ABB RAPID module: MainProgram.mod

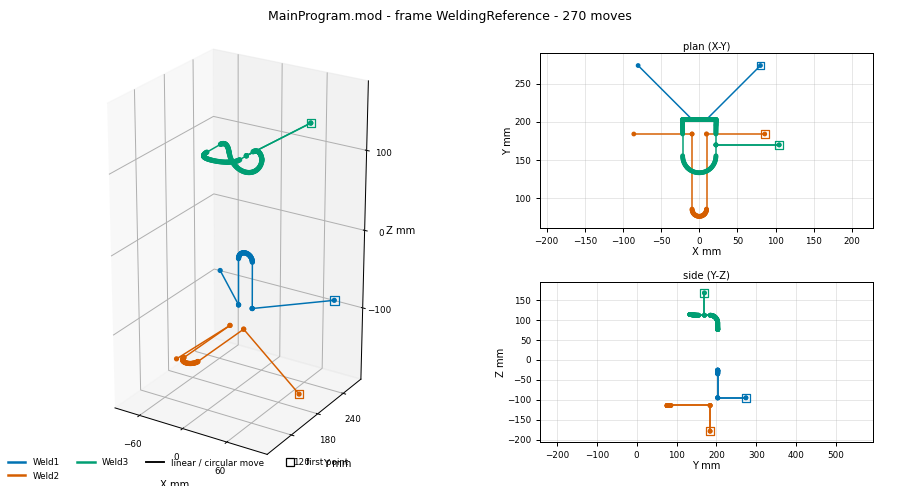
[picture p0: tool path of MainProgram.mod in frame WeldingReference, 270 of 274 moves have a stored position in this frame; points joined in program order, loops and branches not executed]
%%%
  VERSION:1
  LANGUAGE:ENGLISH
%%%
MODULE MOD_MainProgram

    ! -------------------------------
    ! Define customized variables here
    ! ...

	! Tool variables:
	PERS tooldata Weldgun := [TRUE,[[-4.000,0.000,371.300],[0.92387953,0.00000000,0.38268343,0.00000001]],[1,[0,0,20],[1,0,0,0],0,0,0.005]];

	! Reference variables:
	PERS wobjdata WeldingReference := [FALSE, TRUE, "", [[0,0,0],[1,0,0,0]],[[907.213,-302.346,276.168],[0.70442562,0.70442562,-0.06151869,-0.06151869]]];

	PROC GoHome()
		ConfJ \On;
		ConfL \Off;
		MoveAbsJ [[-0.000000,-14.941300,9.781060,0.000000,57.564300,-0.000000],[9E+09,9E+09,9E+09,9E+09,9E+09,9E+09]],v500,z1,Weldgun \WObj:=WeldingReference;
	ENDPROC

	PROC Weld1()
		ConfJ \On;
		ConfL \Off;
		WeldingReference := [FALSE, TRUE, "", [[0,0,0],[1,0,0,0]],[[907.213,-302.346,276.168],[0.70442562,0.70442562,-0.06151869,-0.06151869]]];
		Weldgun := [TRUE,[[-4.000,0.000,371.300],[0.92387953,0.00000000,0.38268343,0.00000001]],[1,[0,0,20],[1,0,0,0],0,0,0.005]];
		! show Weld gun
		MoveAbsJ [[-12.555800,6.650190,11.177100,0.026927,72.173900,-2.607590],[9E+09,9E+09,9E+09,9E+09,9E+09,9E+09]],v1000,z1,Weldgun \WObj:=WeldingReference;
		SetRPM 70.0;
		MoveL [[80.178,273.912,-94.776],[0.27080492,-0.27039115,-0.65336714,0.65319576],[-1,0,-1,0],[9E+09,9E+09,9E+09,9E+09,9E+09,9E+09]],[16.67,500,5000,1000],z1,Weldgun \WObj:=WeldingReference;
		MoveL [[9.468,203.201,-94.776],[0.27080492,-0.27039115,-0.65336714,0.65319576],[-1,0,-1,0],[9E+09,9E+09,9E+09,9E+09,9E+09,9E+09]],[16.67,500,5000,1000],z1,Weldgun \WObj:=WeldingReference;
		GunOn;
		MoveL [[9.468,203.201,-94.776],[0.27080492,-0.27039115,-0.65336714,0.65319576],[-1,0,-1,0],[9E+09,9E+09,9E+09,9E+09,9E+09,9E+09]],[16.67,500,5000,1000],z1,Weldgun \WObj:=WeldingReference;
		MoveL [[9.521,203.201,-94.770],[0.27059813,-0.27059797,-0.65328151,0.65328145],[-1,0,-1,0],[9E+09,9E+09,9E+09,9E+09,9E+09,9E+09]],[16.67,500,5000,1000],z1,Weldgun \WObj:=WeldingReference;
		MoveL [[9.521,203.201,-34.925],[0.26109596,-0.28004323,-0.64928868,0.65713689],[-1,-1,-1,0],[9E+09,9E+09,9E+09,9E+09,9E+09,9E+09]],[16.67,500,5000,1000],z1,Weldgun \WObj:=WeldingReference;
		MoveL [[9.489,203.201,-34.145],[0.23425026,-0.30675221,-0.65944853,0.64510273],[-1,-1,0,0],[9E+09,9E+09,9E+09,9E+09,9E+09,9E+09]],[16.67,500,5000,1000],z1,Weldgun \WObj:=WeldingReference;
		MoveL [[9.394,203.201,-33.370],[0.20701375,-0.33294335,-0.66849979,0.63198265],[-1,-1,0,0],[9E+09,9E+09,9E+09,9E+09,9E+09,9E+09]],[16.67,500,5000,1000],z1,Weldgun \WObj:=WeldingReference;
		MoveL [[9.235,203.201,-32.605],[0.17943264,-0.35858122,-0.67642029,0.61780177],[-1,-1,0,0],[9E+09,9E+09,9E+09,9E+09,9E+09,9E+09]],[16.67,500,5000,1000],z1,Weldgun \WObj:=WeldingReference;
		MoveL [[9.014,203.201,-31.857],[0.15154219,-0.38361099,-0.68321444,0.60257415],[-1,-1,0,0],[9E+09,9E+09,9E+09,9E+09,9E+09,9E+09]],[16.67,500,5000,1000],z1,Weldgun \WObj:=WeldingReference;
		MoveL [[8.732,203.201,-31.128],[0.12340353,-0.40798899,-0.68885701,0.58633828],[-1,-1,0,0],[9E+09,9E+09,9E+09,9E+09,9E+09,9E+09]],[16.67,500,5000,1000],z1,Weldgun \WObj:=WeldingReference;
		MoveL [[8.391,203.201,-30.426],[0.09505233,-0.43169103,-0.69333556,0.56911660],[-1,-1,0,0],[9E+09,9E+09,9E+09,9E+09,9E+09,9E+09]],[16.67,500,5000,1000],z1,Weldgun \WObj:=WeldingReference;
		MoveL [[7.994,203.201,-29.753],[0.06655006,-0.45466761,-0.69664493,0.55093947],[-1,-1,0,0],[9E+09,9E+09,9E+09,9E+09,9E+09,9E+09]],[16.67,500,5000,1000],z1,Weldgun \WObj:=WeldingReference;
		MoveL [[7.544,203.201,-29.116],[0.03792629,-0.47687790,-0.69878733,0.53183205],[-1,-1,0,0],[9E+09,9E+09,9E+09,9E+09,9E+09,9E+09]],[16.67,500,5000,1000],z1,Weldgun \WObj:=WeldingReference;
		MoveL [[7.042,203.201,-28.517],[0.01240330,-0.49395227,-0.70281556,0.51176909],[-1,-1,0,0],[9E+09,9E+09,9E+09,9E+09,9E+09,9E+09]],[16.67,500,5000,1000],z1,Weldgun \WObj:=WeldingReference;
		MoveL [[6.733,203.201,-28.192],[0.00416831,0.50587340,0.70291668,-0.49998286],[-1,-1,0,0],[9E+09,9E+09,9E+09,9E+09,9E+09,9E+09]],[16.67,500,5000,1000],z1,Weldgun \WObj:=WeldingReference;
		MoveL [[6.408,203.201,-27.883],[0.02374061,0.52184249,0.69941540,-0.48778571],[-1,-1,0,0],[9E+09,9E+09,9E+09,9E+09,9E+09,9E+09]],[16.67,500,5000,1000],z1,Weldgun \WObj:=WeldingReference;
		MoveL [[5.809,203.201,-27.381],[0.05240062,0.54140968,0.69785181,-0.46597487],[-1,-1,0,0],[9E+09,9E+09,9E+09,9E+09,9E+09,9E+09]],[16.67,500,5000,1000],z1,Weldgun \WObj:=WeldingReference;
		MoveL [[5.172,203.201,-26.930],[0.08097272,0.56005587,0.69511960,-0.44338425],[-1,-1,0,0],[9E+09,9E+09,9E+09,9E+09,9E+09,9E+09]],[16.67,500,5000,1000],z1,Weldgun \WObj:=WeldingReference;
		MoveL [[4.499,203.201,-26.534],[0.10940637,0.57776774,0.69121158,-0.42004909],[-1,-1,0,0],[9E+09,9E+09,9E+09,9E+09,9E+09,9E+09]],[16.67,500,5000,1000],z1,Weldgun \WObj:=WeldingReference;
		MoveL [[3.797,203.201,-26.193],[0.13765258,0.59450380,0.68614585,-0.39600615],[-1,-1,0,0],[9E+09,9E+09,9E+09,9E+09,9E+09,9E+09]],[16.67,500,5000,1000],z1,Weldgun \WObj:=WeldingReference;
		MoveL [[3.068,203.201,-25.912],[0.16567219,0.61024237,0.67992465,-0.37129428],[-1,-1,0,0],[9E+09,9E+09,9E+09,9E+09,9E+09,9E+09]],[16.67,500,5000,1000],z1,Weldgun \WObj:=WeldingReference;
		MoveL [[2.320,203.201,-25.690],[0.19341081,0.62495524,0.67255736,-0.34596213],[-1,-1,0,0],[9E+09,9E+09,9E+09,9E+09,9E+09,9E+09]],[16.67,500,5000,1000],z1,Weldgun \WObj:=WeldingReference;
		MoveL [[1.555,203.201,-25.531],[0.22082406,0.63861348,0.66406224,-0.32004826],[-1,-1,0,0],[9E+09,9E+09,9E+09,9E+09,9E+09,9E+09]],[16.67,500,5000,1000],z1,Weldgun \WObj:=WeldingReference;
		MoveL [[0.780,203.201,-25.436],[0.24786932,0.65119902,0.65444982,-0.29359169],[-1,-1,0,0],[9E+09,9E+09,9E+09,9E+09,9E+09,9E+09]],[16.67,500,5000,1000],z1,Weldgun \WObj:=WeldingReference;
		MoveL [[0.000,203.201,-25.404],[0.27449275,0.66268723,0.64373837,-0.26664635],[-1,-1,0,0],[9E+09,9E+09,9E+09,9E+09,9E+09,9E+09]],[16.67,500,5000,1000],z1,Weldgun \WObj:=WeldingReference;
		MoveL [[-0.780,203.201,-25.436],[0.30065949,0.67306272,0.63194229,-0.23924755],[-1,-1,0,0],[9E+09,9E+09,9E+09,9E+09,9E+09,9E+09]],[16.67,500,5000,1000],z1,Weldgun \WObj:=WeldingReference;
		MoveL [[-1.555,203.201,-25.531],[0.32631571,0.68230801,0.61908153,-0.21145189],[-1,0,1,0],[9E+09,9E+09,9E+09,9E+09,9E+09,9E+09]],[16.67,500,5000,1000],z1,Weldgun \WObj:=WeldingReference;
		MoveL [[-2.320,203.201,-25.690],[0.35142970,0.69040355,0.60518073,-0.18329319],[-1,0,1,0],[9E+09,9E+09,9E+09,9E+09,9E+09,9E+09]],[16.67,500,5000,1000],z1,Weldgun \WObj:=WeldingReference;
		MoveL [[-3.068,203.201,-25.912],[0.37594474,0.69734095,0.59026085,-0.15483308],[-1,0,1,0],[9E+09,9E+09,9E+09,9E+09,9E+09,9E+09]],[16.67,500,5000,1000],z1,Weldgun \WObj:=WeldingReference;
		MoveL [[-3.797,203.201,-26.193],[0.39983154,0.70309811,0.57435509,-0.12611111],[-1,0,1,0],[9E+09,9E+09,9E+09,9E+09,9E+09,9E+09]],[16.67,500,5000,1000],z1,Weldgun \WObj:=WeldingReference;
		MoveL [[-4.499,203.201,-26.534],[0.42304339,0.70768163,0.55747448,-0.09717615],[-1,0,1,0],[9E+09,9E+09,9E+09,9E+09,9E+09,9E+09]],[16.67,500,5000,1000],z1,Weldgun \WObj:=WeldingReference;
		MoveL [[-5.172,203.201,-26.930],[0.44554480,0.71107104,0.53966024,-0.06807809],[-1,0,1,0],[9E+09,9E+09,9E+09,9E+09,9E+09,9E+09]],[16.67,500,5000,1000],z1,Weldgun \WObj:=WeldingReference;
		MoveL [[-5.809,203.201,-27.381],[0.46730140,0.71326404,0.52093536,-0.03886082],[-1,0,1,0],[9E+09,9E+09,9E+09,9E+09,9E+09,9E+09]],[16.67,500,5000,1000],z1,Weldgun \WObj:=WeldingReference;
		MoveL [[-6.408,203.201,-27.883],[0.48819595,0.71113015,0.50576611,-0.01261974],[-1,0,1,0],[9E+09,9E+09,9E+09,9E+09,9E+09,9E+09]],[16.67,500,5000,1000],z1,Weldgun \WObj:=WeldingReference;
		MoveL [[-6.731,203.201,-28.191],[0.49992546,0.71126987,0.49411825,0.00410579],[-1,0,1,0],[9E+09,9E+09,9E+09,9E+09,9E+09,9E+09]],[16.67,500,5000,1000],z1,Weldgun \WObj:=WeldingReference;
		MoveL [[-7.042,203.201,-28.517],[0.51134749,0.71391546,0.47777457,0.02408169],[-1,0,1,0],[9E+09,9E+09,9E+09,9E+09,9E+09,9E+09]],[16.67,500,5000,1000],z1,Weldgun \WObj:=WeldingReference;
		MoveL [[-7.544,203.201,-29.116],[0.53050914,0.71232829,0.45640294,0.05333687],[-1,0,1,0],[9E+09,9E+09,9E+09,9E+09,9E+09,9E+09]],[16.67,500,5000,1000],z1,Weldgun \WObj:=WeldingReference;
		MoveL [[-7.994,203.201,-29.753],[0.54878026,0.70953905,0.43426730,0.08250137],[-1,0,1,0],[9E+09,9E+09,9E+09,9E+09,9E+09,9E+09]],[16.67,500,5000,1000],z1,Weldgun \WObj:=WeldingReference;
		MoveL [[-8.391,203.201,-30.426],[0.56612441,0.70556165,0.41139698,0.11152774],[-1,0,1,0],[9E+09,9E+09,9E+09,9E+09,9E+09,9E+09]],[16.67,500,5000,1000],z1,Weldgun \WObj:=WeldingReference;
		MoveL [[-8.732,203.201,-31.128],[0.58251728,0.70039316,0.38784300,0.14035973],[-1,0,1,0],[9E+09,9E+09,9E+09,9E+09,9E+09,9E+09]],[16.67,500,5000,1000],z1,Weldgun \WObj:=WeldingReference;
		MoveL [[-9.014,203.201,-31.857],[0.59792965,0.69404912,0.36363243,0.16895976],[-1,0,1,0],[9E+09,9E+09,9E+09,9E+09,9E+09,9E+09]],[16.67,500,5000,1000],z1,Weldgun \WObj:=WeldingReference;
		MoveL [[-9.235,203.201,-32.605],[0.61233261,0.68654186,0.33880881,0.19727554],[-1,0,1,0],[9E+09,9E+09,9E+09,9E+09,9E+09,9E+09]],[16.67,500,5000,1000],z1,Weldgun \WObj:=WeldingReference;
		MoveL [[-9.394,203.201,-33.370],[0.62571166,0.67787385,0.31341661,0.22525981],[-1,0,1,0],[9E+09,9E+09,9E+09,9E+09,9E+09,9E+09]],[16.67,500,5000,1000],z1,Weldgun \WObj:=WeldingReference;
		MoveL [[-9.489,203.201,-34.145],[0.63803534,0.66806855,0.28749564,0.25286671],[-1,0,1,0],[9E+09,9E+09,9E+09,9E+09,9E+09,9E+09]],[16.67,500,5000,1000],z1,Weldgun \WObj:=WeldingReference;
		MoveL [[-9.521,203.201,-34.925],[0.65328148,0.65328148,0.27059805,0.27059805],[-1,0,1,0],[9E+09,9E+09,9E+09,9E+09,9E+09,9E+09]],[16.67,500,5000,1000],z1,Weldgun \WObj:=WeldingReference;
		MoveL [[-9.521,203.201,-94.770],[0.65328148,0.65328148,0.27059805,0.27059805],[-1,0,1,0],[9E+09,9E+09,9E+09,9E+09,9E+09,9E+09]],[16.67,500,5000,1000],z1,Weldgun \WObj:=WeldingReference;
		MoveL [[-9.470,203.201,-94.776],[0.65328148,0.65328148,0.27059805,0.27059805],[-1,0,1,0],[9E+09,9E+09,9E+09,9E+09,9E+09,9E+09]],[16.67,500,5000,1000],z1,Weldgun \WObj:=WeldingReference;
		GunOff;
		MoveL [[-9.470,203.201,-94.776],[0.65328148,0.65328148,0.27059805,0.27059805],[-1,0,1,0],[9E+09,9E+09,9E+09,9E+09,9E+09,9E+09]],v1000,z1,Weldgun \WObj:=WeldingReference;
		MoveL [[-80.181,273.912,-94.776],[0.65328148,0.65328148,0.27059805,0.27059805],[-1,0,1,0],[9E+09,9E+09,9E+09,9E+09,9E+09,9E+09]],v1000,z1,Weldgun \WObj:=WeldingReference;
	ENDPROC

	PROC Weld2()
		ConfJ \On;
		ConfL \Off;
		WeldingReference := [FALSE, TRUE, "", [[0,0,0],[1,0,0,0]],[[907.213,-302.346,276.168],[0.70442562,0.70442562,-0.06151869,-0.06151869]]];
		Weldgun := [TRUE,[[-4.000,0.000,371.300],[0.92387953,0.00000000,0.38268343,0.00000001]],[1,[0,0,20],[1,0,0,0],0,0,0.005]];
		! show Weld gun
		MoveAbsJ [[14.847000,37.704900,12.622700,-66.388600,108.377000,54.200400],[9E+09,9E+09,9E+09,9E+09,9E+09,9E+09]],v1000,z1,Weldgun \WObj:=WeldingReference;
		SetRPM 70.0;
		MoveL [[85.827,184.150,-178.501],[0.00000000,-0.42074767,0.00000000,0.90717771],[0,-1,0,0],[9E+09,9E+09,9E+09,9E+09,9E+09,9E+09]],[16.67,500,5000,1000],z1,Weldgun \WObj:=WeldingReference;
		MoveL [[9.489,184.150,-113.907],[0.00000000,-0.42074767,0.00000000,0.90717771],[0,-1,0,0],[9E+09,9E+09,9E+09,9E+09,9E+09,9E+09]],[16.67,500,5000,1000],z1,Weldgun \WObj:=WeldingReference;
		GunOn;
		MoveL [[9.489,184.150,-113.907],[0.00000000,-0.42074767,0.00000000,0.90717771],[0,-1,0,0],[9E+09,9E+09,9E+09,9E+09,9E+09,9E+09]],[16.67,500,5000,1000],z1,Weldgun \WObj:=WeldingReference;
		MoveL [[9.489,85.725,-113.907],[0.01312106,-0.42070385,-0.00608599,0.90708273],[0,-1,0,0],[9E+09,9E+09,9E+09,9E+09,9E+09,9E+09]],[16.67,500,5000,1000],z1,Weldgun \WObj:=WeldingReference;
		MoveL [[9.457,84.942,-113.910],[0.05153547,-0.42042592,0.00808679,0.90582600],[0,-1,0,0],[9E+09,9E+09,9E+09,9E+09,9E+09,9E+09]],[16.67,500,5000,1000],z1,Weldgun \WObj:=WeldingReference;
		MoveL [[9.361,84.163,-113.917],[0.08985371,-0.41918442,0.02228324,0.90316897],[0,-1,0,0],[9E+09,9E+09,9E+09,9E+09,9E+09,9E+09]],[16.67,500,5000,1000],z1,Weldgun \WObj:=WeldingReference;
		MoveL [[9.202,83.396,-113.930],[0.12804465,-0.41698615,0.03650971,0.89910742],[0,-1,0,0],[9E+09,9E+09,9E+09,9E+09,9E+09,9E+09]],[16.67,500,5000,1000],z1,Weldgun \WObj:=WeldingReference;
		MoveL [[8.981,82.644,-113.948],[0.16597915,-0.41384219,0.05079357,0.89364735],[0,-1,0,0],[9E+09,9E+09,9E+09,9E+09,9E+09,9E+09]],[16.67,500,5000,1000],z1,Weldgun \WObj:=WeldingReference;
		MoveL [[8.700,81.913,-113.970],[0.20363787,-0.40977344,0.06511381,0.88677931],[0,-1,0,0],[9E+09,9E+09,9E+09,9E+09,9E+09,9E+09]],[16.67,500,5000,1000],z1,Weldgun \WObj:=WeldingReference;
		MoveL [[8.360,81.208,-113.995],[0.24095022,-0.40479903,0.07948489,0.87850037],[0,-1,0,0],[9E+09,9E+09,9E+09,9E+09,9E+09,9E+09]],[16.67,500,5000,1000],z1,Weldgun \WObj:=WeldingReference;
		MoveL [[7.963,80.534,-114.024],[0.27783978,-0.39894829,0.09389601,0.86880887],[0,-1,0,0],[9E+09,9E+09,9E+09,9E+09,9E+09,9E+09]],[16.67,500,5000,1000],z1,Weldgun \WObj:=WeldingReference;
		MoveL [[7.512,79.895,-114.054],[0.31416482,-0.39224451,0.10838187,0.85772844],[0,-1,0,0],[9E+09,9E+09,9E+09,9E+09,9E+09,9E+09]],[16.67,500,5000,1000],z1,Weldgun \WObj:=WeldingReference;
		MoveL [[7.009,79.295,-114.086],[0.34473394,-0.38397214,0.12525349,0.84736974],[0,-1,0,0],[9E+09,9E+09,9E+09,9E+09,9E+09,9E+09]],[16.67,500,5000,1000],z1,Weldgun \WObj:=WeldingReference;
		MoveL [[6.707,78.978,-114.104],[0.36453651,-0.37938408,0.13335075,0.83988001],[0,-1,0,0],[9E+09,9E+09,9E+09,9E+09,9E+09,9E+09]],[16.67,500,5000,1000],z1,Weldgun \WObj:=WeldingReference;
		MoveL [[6.391,78.676,-114.123],[0.38912980,-0.37541067,0.13918584,0.82962168],[0,-1,0,0],[9E+09,9E+09,9E+09,9E+09,9E+09,9E+09]],[16.67,500,5000,1000],z1,Weldgun \WObj:=WeldingReference;
		MoveL [[5.795,78.176,-114.154],[0.42321516,-0.36636835,0.15366636,0.81427871],[0,-1,0,0],[9E+09,9E+09,9E+09,9E+09,9E+09,9E+09]],[16.67,500,5000,1000],z1,Weldgun \WObj:=WeldingReference;
		MoveL [[5.160,77.727,-114.185],[0.45649477,-0.35666115,0.16813439,0.79758145],[0,-1,0,0],[9E+09,9E+09,9E+09,9E+09,9E+09,9E+09]],[16.67,500,5000,1000],z1,Weldgun \WObj:=WeldingReference;
		MoveL [[4.490,77.331,-114.213],[0.48887672,-0.34632893,0.18258429,0.77956321],[0,-1,0,0],[9E+09,9E+09,9E+09,9E+09,9E+09,9E+09]],[16.67,500,5000,1000],z1,Weldgun \WObj:=WeldingReference;
		MoveL [[3.790,76.991,-114.239],[0.52034210,-0.33543360,0.19697026,0.76021781],[0,-1,-1,0],[9E+09,9E+09,9E+09,9E+09,9E+09,9E+09]],[16.67,500,5000,1000],z1,Weldgun \WObj:=WeldingReference;
		MoveL [[3.063,76.710,-114.260],[0.55080992,-0.32401460,0.21128182,0.73958297],[0,-1,-1,0],[9E+09,9E+09,9E+09,9E+09,9E+09,9E+09]],[16.67,500,5000,1000],z1,Weldgun \WObj:=WeldingReference;
		MoveL [[2.316,76.490,-114.278],[0.58023779,-0.31212946,0.22547321,0.71767759],[0,-1,-1,0],[9E+09,9E+09,9E+09,9E+09,9E+09,9E+09]],[16.67,500,5000,1000],z1,Weldgun \WObj:=WeldingReference;
		MoveL [[1.553,76.331,-114.291],[0.60858630,-0.29982600,0.23951509,0.69452113],[0,-1,-1,0],[9E+09,9E+09,9E+09,9E+09,9E+09,9E+09]],[16.67,500,5000,1000],z1,Weldgun \WObj:=WeldingReference;
		MoveL [[0.779,76.236,-114.299],[0.63581862,-0.28715637,0.25336406,0.67013622],[0,-1,-1,0],[9E+09,9E+09,9E+09,9E+09,9E+09,9E+09]],[16.67,500,5000,1000],z1,Weldgun \WObj:=WeldingReference;
		MoveL [[0.000,76.204,-114.301],[0.66190027,-0.27416831,0.26698017,0.64454741],[0,-1,-1,0],[9E+09,9E+09,9E+09,9E+09,9E+09,9E+09]],[16.67,500,5000,1000],z1,Weldgun \WObj:=WeldingReference;
		MoveL [[-0.779,76.236,-114.299],[0.68679970,-0.26090700,0.28032057,0.61778159],[0,-1,-1,0],[9E+09,9E+09,9E+09,9E+09,9E+09,9E+09]],[16.67,500,5000,1000],z1,Weldgun \WObj:=WeldingReference;
		MoveL [[-1.553,76.331,-114.291],[0.71048565,-0.24741615,0.29333969,0.58987051],[0,-1,-1,0],[9E+09,9E+09,9E+09,9E+09,9E+09,9E+09]],[16.67,500,5000,1000],z1,Weldgun \WObj:=WeldingReference;
		MoveL [[-2.316,76.490,-114.278],[0.73293327,-0.23373805,0.30598954,0.56084377],[0,-1,-1,0],[9E+09,9E+09,9E+09,9E+09,9E+09,9E+09]],[16.67,500,5000,1000],z1,Weldgun \WObj:=WeldingReference;
		MoveL [[-3.063,76.710,-114.260],[0.75411156,-0.21990803,0.31822287,0.53074516],[0,-1,-1,0],[9E+09,9E+09,9E+09,9E+09,9E+09,9E+09]],[16.67,500,5000,1000],z1,Weldgun \WObj:=WeldingReference;
		MoveL [[-3.790,76.991,-114.239],[0.77400420,-0.20596628,0.32998612,0.49960440],[0,-1,-1,0],[9E+09,9E+09,9E+09,9E+09,9E+09,9E+09]],[16.67,500,5000,1000],z1,Weldgun \WObj:=WeldingReference;
		MoveL [[-4.490,77.331,-114.213],[0.79256096,-0.19192832,0.34123966,0.46751058],[0,-1,-1,0],[9E+09,9E+09,9E+09,9E+09,9E+09,9E+09]],[16.67,500,5000,1000],z1,Weldgun \WObj:=WeldingReference;
		MoveL [[-5.160,77.727,-114.185],[0.80978515,-0.17783865,0.35192282,0.43447872],[0,-1,-1,0],[9E+09,9E+09,9E+09,9E+09,9E+09,9E+09]],[16.67,500,5000,1000],z1,Weldgun \WObj:=WeldingReference;
		MoveL [[-5.795,78.176,-114.154],[0.82563537,-0.16370520,0.36199413,0.40060840],[0,-1,-1,0],[9E+09,9E+09,9E+09,9E+09,9E+09,9E+09]],[16.67,500,5000,1000],z1,Weldgun \WObj:=WeldingReference;
		MoveL [[-6.391,78.676,-114.123],[0.83783925,-0.14727053,0.37231303,0.37110616],[0,-1,-1,0],[9E+09,9E+09,9E+09,9E+09,9E+09,9E+09]],[16.67,500,5000,1000],z1,Weldgun \WObj:=WeldingReference;
		MoveL [[-6.706,78.977,-114.105],[0.84546949,-0.13933620,0.37721701,0.35138881],[0,-1,-1,0],[9E+09,9E+09,9E+09,9E+09,9E+09,9E+09]],[16.67,500,5000,1000],z1,Weldgun \WObj:=WeldingReference;
		MoveL [[-7.009,79.295,-114.086],[0.85473835,-0.13366178,0.38112708,0.32603532],[0,-1,-1,0],[9E+09,9E+09,9E+09,9E+09,9E+09,9E+09]],[16.67,500,5000,1000],z1,Weldgun \WObj:=WeldingReference;
		MoveL [[-7.512,79.895,-114.054],[0.86625855,-0.11941761,0.38902742,0.28981584],[0,-1,-1,0],[9E+09,9E+09,9E+09,9E+09,9E+09,9E+09]],[16.67,500,5000,1000],z1,Weldgun \WObj:=WeldingReference;
		MoveL [[-7.963,80.534,-114.024],[0.87636361,-0.10521269,0.39611442,0.25300292],[0,-1,-1,0],[9E+09,9E+09,9E+09,9E+09,9E+09,9E+09]],[16.67,500,5000,1000],z1,Weldgun \WObj:=WeldingReference;
		MoveL [[-8.360,81.208,-113.995],[0.88502630,-0.09101818,0.40236240,0.21575135],[0,-1,-1,0],[9E+09,9E+09,9E+09,9E+09,9E+09,9E+09]],[16.67,500,5000,1000],z1,Weldgun \WObj:=WeldingReference;
		MoveL [[-8.700,81.913,-113.970],[0.89225386,-0.07683939,0.40773709,0.17812700],[0,-1,-2,0],[9E+09,9E+09,9E+09,9E+09,9E+09,9E+09]],[16.67,500,5000,1000],z1,Weldgun \WObj:=WeldingReference;
		MoveL [[-8.981,82.644,-113.948],[0.89804934,-0.06266887,0.41221168,0.14021956],[0,-1,-2,0],[9E+09,9E+09,9E+09,9E+09,9E+09,9E+09]],[16.67,500,5000,1000],z1,Weldgun \WObj:=WeldingReference;
		MoveL [[-9.202,83.396,-113.930],[0.90242768,-0.04852727,0.41575907,0.10204796],[0,-1,-2,0],[9E+09,9E+09,9E+09,9E+09,9E+09,9E+09]],[16.67,500,5000,1000],z1,Weldgun \WObj:=WeldingReference;
		MoveL [[-9.361,84.163,-113.917],[0.90538716,-0.03438326,0.41836580,0.06373333],[0,-1,-2,0],[9E+09,9E+09,9E+09,9E+09,9E+09,9E+09]],[16.67,500,5000,1000],z1,Weldgun \WObj:=WeldingReference;
		MoveL [[-9.457,84.942,-113.910],[0.90693713,-0.02023844,0.42001684,0.02532396],[0,-1,-2,0],[9E+09,9E+09,9E+09,9E+09,9E+09,9E+09]],[16.67,500,5000,1000],z1,Weldgun \WObj:=WeldingReference;
		MoveL [[-9.489,85.725,-113.907],[0.90717771,0.00000000,0.42074767,0.00000000],[0,-1,-2,0],[9E+09,9E+09,9E+09,9E+09,9E+09,9E+09]],[16.67,500,5000,1000],z1,Weldgun \WObj:=WeldingReference;
		MoveL [[-9.489,184.150,-113.907],[0.90717771,0.00000000,0.42074767,0.00000000],[0,-1,-2,0],[9E+09,9E+09,9E+09,9E+09,9E+09,9E+09]],[16.67,500,5000,1000],z1,Weldgun \WObj:=WeldingReference;
		GunOff;
		MoveL [[-9.489,184.150,-113.907],[0.90717771,0.00000000,0.42074767,0.00000000],[0,-1,-2,0],[9E+09,9E+09,9E+09,9E+09,9E+09,9E+09]],v1000,z1,Weldgun \WObj:=WeldingReference;
		MoveL [[-85.827,184.150,-178.501],[0.90717771,0.00000000,0.42074767,0.00000000],[0,-1,-2,0],[9E+09,9E+09,9E+09,9E+09,9E+09,9E+09]],v1000,z1,Weldgun \WObj:=WeldingReference;
	ENDPROC

	PROC Weld3()
		ConfJ \On;
		ConfL \Off;
		WeldingReference := [FALSE, TRUE, "", [[0,0,0],[1,0,0,0]],[[907.213,-302.346,276.168],[0.70442562,0.70442562,-0.06151869,-0.06151869]]];
		Weldgun := [TRUE,[[-4.000,0.000,371.300],[0.92387953,0.00000000,0.38268343,0.00000001]],[1,[0,0,20],[1,0,0,0],0,0,0.005]];
		! show Weld gun
		MoveAbsJ [[-42.441800,44.926500,-10.306700,45.964800,113.439000,-33.438500],[9E+09,9E+09,9E+09,9E+09,9E+09,9E+09]],v1000,z1,Weldgun \WObj:=WeldingReference;
		SetRPM 70.0;
		MoveL [[104.720,169.863,168.115],[0.45836971,-0.19110070,-0.86200423,0.10161911],[-1,0,-1,0],[9E+09,9E+09,9E+09,9E+09,9E+09,9E+09]],[16.67,500,5000,1000],z1,Weldgun \WObj:=WeldingReference;
		MoveL [[21.813,169.863,112.201],[0.46949853,-0.00000000,-0.88293325,0.00000000],[-1,0,-1,0],[9E+09,9E+09,9E+09,9E+09,9E+09,9E+09]],[16.67,500,5000,1000],z1,Weldgun \WObj:=WeldingReference;
		GunOn;
		MoveL [[21.813,169.863,112.201],[0.46949853,-0.00000000,-0.88293325,0.00000000],[-1,0,-1,0],[9E+09,9E+09,9E+09,9E+09,9E+09,9E+09]],[16.67,500,5000,1000],z1,Weldgun \WObj:=WeldingReference;
		MoveL [[21.813,155.575,112.201],[0.46947851,-0.00826181,-0.88289433,0.00439085],[-1,0,-1,0],[9E+09,9E+09,9E+09,9E+09,9E+09,9E+09]],[16.67,500,5000,1000],z1,Weldgun \WObj:=WeldingReference;
		MoveL [[21.782,154.355,112.207],[0.46925544,-0.03372123,-0.88241081,-0.00365648],[-1,0,-1,0],[9E+09,9E+09,9E+09,9E+09,9E+09,9E+09]],[16.67,500,5000,1000],z1,Weldgun \WObj:=WeldingReference;
		MoveL [[21.686,153.139,112.225],[0.46843794,-0.05917155,-0.88143470,-0.01172583],[-1,0,-1,0],[9E+09,9E+09,9E+09,9E+09,9E+09,9E+09]],[16.67,500,5000,1000],z1,Weldgun \WObj:=WeldingReference;
		MoveL [[21.528,151.930,112.256],[0.46702608,-0.08461970,-0.87996163,-0.01984127],[-1,0,-1,0],[9E+09,9E+09,9E+09,9E+09,9E+09,9E+09]],[16.67,500,5000,1000],z1,Weldgun \WObj:=WeldingReference;
		MoveL [[21.307,150.732,112.298],[0.46502371,-0.10999279,-0.87799155,-0.02802444],[-1,0,-1,0],[9E+09,9E+09,9E+09,9E+09,9E+09,9E+09]],[16.67,500,5000,1000],z1,Weldgun \WObj:=WeldingReference;
		MoveL [[21.026,149.557,112.351],[0.46245601,-0.13521188,-0.87552324,-0.03621095],[-1,0,-1,0],[9E+09,9E+09,9E+09,9E+09,9E+09,9E+09]],[16.67,500,5000,1000],z1,Weldgun \WObj:=WeldingReference;
		MoveL [[20.685,148.403,112.414],[0.45932769,-0.16034081,-0.87254456,-0.04443977],[-1,0,-1,0],[9E+09,9E+09,9E+09,9E+09,9E+09,9E+09]],[16.67,500,5000,1000],z1,Weldgun \WObj:=WeldingReference;
		MoveL [[20.284,147.270,112.487],[0.45564189,-0.18539904,-0.86904213,-0.05275829],[-1,0,-1,0],[9E+09,9E+09,9E+09,9E+09,9E+09,9E+09]],[16.67,500,5000,1000],z1,Weldgun \WObj:=WeldingReference;
		MoveL [[19.824,146.161,112.569],[0.45140558,-0.21040952,-0.86499545,-0.06118584],[-1,0,-1,0],[9E+09,9E+09,9E+09,9E+09,9E+09,9E+09]],[16.67,500,5000,1000],z1,Weldgun \WObj:=WeldingReference;
		MoveL [[19.306,145.081,112.659],[0.44663266,-0.23530443,-0.86040042,-0.06972955],[-1,0,-1,0],[9E+09,9E+09,9E+09,9E+09,9E+09,9E+09]],[16.67,500,5000,1000],z1,Weldgun \WObj:=WeldingReference;
		MoveL [[18.731,144.031,112.756],[0.44133315,-0.26008182,-0.85523924,-0.07841129],[-1,0,-1,0],[9E+09,9E+09,9E+09,9E+09,9E+09,9E+09]],[16.67,500,5000,1000],z1,Weldgun \WObj:=WeldingReference;
		MoveL [[18.101,143.016,112.859],[0.43552760,-0.28469939,-0.84950197,-0.08722601],[-1,0,-1,0],[9E+09,9E+09,9E+09,9E+09,9E+09,9E+09]],[16.67,500,5000,1000],z1,Weldgun \WObj:=WeldingReference;
		MoveL [[17.416,142.038,112.967],[0.42922926,-0.30911875,-0.84318181,-0.09618877],[-1,0,-1,0],[9E+09,9E+09,9E+09,9E+09,9E+09,9E+09]],[16.67,500,5000,1000],z1,Weldgun \WObj:=WeldingReference;
		MoveL [[16.680,141.100,113.078],[0.42245731,-0.33330391,-0.83626980,-0.10531455],[-1,0,-1,0],[9E+09,9E+09,9E+09,9E+09,9E+09,9E+09]],[16.67,500,5000,1000],z1,Weldgun \WObj:=WeldingReference;
		MoveL [[15.892,140.204,113.191],[0.41479773,-0.35408689,-0.83010196,-0.11617253],[-1,0,-1,0],[9E+09,9E+09,9E+09,9E+09,9E+09,9E+09]],[16.67,500,5000,1000],z1,Weldgun \WObj:=WeldingReference;
		MoveL [[15.420,139.713,113.257],[0.41045549,-0.36765270,-0.82558355,-0.12153015],[-1,0,-1,0],[9E+09,9E+09,9E+09,9E+09,9E+09,9E+09]],[16.67,500,5000,1000],z1,Weldgun \WObj:=WeldingReference;
		MoveL [[14.932,139.236,113.322],[0.40642995,-0.38404845,-0.81949606,-0.12548980],[-1,0,-1,0],[9E+09,9E+09,9E+09,9E+09,9E+09,9E+09]],[16.67,500,5000,1000],z1,Weldgun \WObj:=WeldingReference;
		MoveL [[14.061,138.456,113.433],[0.39847196,-0.40677858,-0.81088757,-0.13495418],[-1,0,-1,0],[9E+09,9E+09,9E+09,9E+09,9E+09,9E+09]],[16.67,500,5000,1000],z1,Weldgun \WObj:=WeldingReference;
		MoveL [[13.150,137.727,113.542],[0.39018874,-0.42907413,-0.80172291,-0.14452859],[-1,0,-1,0],[9E+09,9E+09,9E+09,9E+09,9E+09,9E+09]],[16.67,500,5000,1000],z1,Weldgun \WObj:=WeldingReference;
		MoveL [[12.201,137.049,113.648],[0.38157390,-0.45094718,-0.79199289,-0.15425712],[-1,0,-1,0],[9E+09,9E+09,9E+09,9E+09,9E+09,9E+09]],[16.67,500,5000,1000],z1,Weldgun \WObj:=WeldingReference;
		MoveL [[11.214,136.423,113.750],[0.37264854,-0.47238051,-0.78169507,-0.16414184],[-1,0,0,0],[9E+09,9E+09,9E+09,9E+09,9E+09,9E+09]],[16.67,500,5000,1000],z1,Weldgun \WObj:=WeldingReference;
		MoveL [[10.194,135.851,113.846],[0.36344534,-0.49334907,-0.77083132,-0.17416445],[-1,0,0,0],[9E+09,9E+09,9E+09,9E+09,9E+09,9E+09]],[16.67,500,5000,1000],z1,Weldgun \WObj:=WeldingReference;
		MoveL [[9.142,135.335,113.935],[0.35399626,-0.51381596,-0.75941325,-0.18431313],[-1,0,0,0],[9E+09,9E+09,9E+09,9E+09,9E+09,9E+09]],[16.67,500,5000,1000],z1,Weldgun \WObj:=WeldingReference;
		MoveL [[8.063,134.876,114.017],[0.34431971,-0.53375533,-0.74745252,-0.19458650],[-1,0,0,0],[9E+09,9E+09,9E+09,9E+09,9E+09,9E+09]],[16.67,500,5000,1000],z1,Weldgun \WObj:=WeldingReference;
		MoveL [[6.958,134.475,114.089],[0.33445023,-0.55318165,-0.73493068,-0.20496340],[-1,0,0,0],[9E+09,9E+09,9E+09,9E+09,9E+09,9E+09]],[16.67,500,5000,1000],z1,Weldgun \WObj:=WeldingReference;
		MoveL [[5.832,134.135,114.153],[0.32440973,-0.57206047,-0.72186741,-0.21543582],[-1,0,0,0],[9E+09,9E+09,9E+09,9E+09,9E+09,9E+09]],[16.67,500,5000,1000],z1,Weldgun \WObj:=WeldingReference;
		MoveL [[4.688,133.854,114.205],[0.31423551,-0.59038635,-0.70826209,-0.22597526],[-1,0,0,0],[9E+09,9E+09,9E+09,9E+09,9E+09,9E+09]],[16.67,500,5000,1000],z1,Weldgun \WObj:=WeldingReference;
		MoveL [[3.529,133.636,114.247],[0.30394438,-0.60817718,-0.69409665,-0.23657592],[-1,0,0,0],[9E+09,9E+09,9E+09,9E+09,9E+09,9E+09]],[16.67,500,5000,1000],z1,Weldgun \WObj:=WeldingReference;
		MoveL [[2.359,133.479,114.277],[0.29355812,-0.62539969,-0.67939583,-0.24722493],[-1,0,0,0],[9E+09,9E+09,9E+09,9E+09,9E+09,9E+09]],[16.67,500,5000,1000],z1,Weldgun \WObj:=WeldingReference;
		MoveL [[1.181,133.385,114.295],[0.28312229,-0.64208469,-0.66412935,-0.25787831],[-1,0,0,0],[9E+09,9E+09,9E+09,9E+09,9E+09,9E+09]],[16.67,500,5000,1000],z1,Weldgun \WObj:=WeldingReference;
		MoveL [[0.000,133.354,114.301],[0.27264144,-0.65820844,-0.64831720,-0.26853883],[-1,0,0,0],[9E+09,9E+09,9E+09,9E+09,9E+09,9E+09]],[16.67,500,5000,1000],z1,Weldgun \WObj:=WeldingReference;
		MoveL [[-1.181,133.385,114.295],[0.26214756,-0.67379835,-0.63193050,-0.27917429],[-1,0,0,0],[9E+09,9E+09,9E+09,9E+09,9E+09,9E+09]],[16.67,500,5000,1000],z1,Weldgun \WObj:=WeldingReference;
		MoveL [[-2.359,133.479,114.277],[0.25165693,-0.68882873,-0.61499449,-0.28976809],[-1,0,0,0],[9E+09,9E+09,9E+09,9E+09,9E+09,9E+09]],[16.67,500,5000,1000],z1,Weldgun \WObj:=WeldingReference;
		MoveL [[-3.529,133.636,114.247],[0.24120568,-0.70332566,-0.59748039,-0.30028322],[-1,0,0,0],[9E+09,9E+09,9E+09,9E+09,9E+09,9E+09]],[16.67,500,5000,1000],z1,Weldgun \WObj:=WeldingReference;
		MoveL [[-4.688,133.854,114.205],[0.23079289,-0.71727319,-0.57940571,-0.31071344],[-1,0,0,0],[9E+09,9E+09,9E+09,9E+09,9E+09,9E+09]],[16.67,500,5000,1000],z1,Weldgun \WObj:=WeldingReference;
		MoveL [[-5.832,134.135,114.153],[0.22044668,-0.73067656,-0.56076483,-0.32102621],[-1,0,0,0],[9E+09,9E+09,9E+09,9E+09,9E+09,9E+09]],[16.67,500,5000,1000],z1,Weldgun \WObj:=WeldingReference;
		MoveL [[-6.958,134.475,114.089],[0.21019099,-0.74353520,-0.54156122,-0.33118968],[-1,0,0,0],[9E+09,9E+09,9E+09,9E+09,9E+09,9E+09]],[16.67,500,5000,1000],z1,Weldgun \WObj:=WeldingReference;
		MoveL [[-8.063,134.876,114.017],[0.20002611,-0.75583225,-0.52182136,-0.34118855],[-1,0,0,0],[9E+09,9E+09,9E+09,9E+09,9E+09,9E+09]],[16.67,500,5000,1000],z1,Weldgun \WObj:=WeldingReference;
		MoveL [[-9.142,135.335,113.935],[0.18997719,-0.76757995,-0.50153408,-0.35098898],[-1,0,0,0],[9E+09,9E+09,9E+09,9E+09,9E+09,9E+09]],[16.67,500,5000,1000],z1,Weldgun \WObj:=WeldingReference;
		MoveL [[-10.194,135.851,113.846],[0.18005715,-0.77876358,-0.48072993,-0.36056267],[-1,0,0,0],[9E+09,9E+09,9E+09,9E+09,9E+09,9E+09]],[16.67,500,5000,1000],z1,Weldgun \WObj:=WeldingReference;
		MoveL [[-11.214,136.423,113.750],[0.17026124,-0.78937111,-0.45943870,-0.36989247],[-1,0,0,0],[9E+09,9E+09,9E+09,9E+09,9E+09,9E+09]],[16.67,500,5000,1000],z1,Weldgun \WObj:=WeldingReference;
		MoveL [[-12.201,137.049,113.648],[0.16060372,-0.79940258,-0.43767835,-0.37894541],[-1,0,0,0],[9E+09,9E+09,9E+09,9E+09,9E+09,9E+09]],[16.67,500,5000,1000],z1,Weldgun \WObj:=WeldingReference;
		MoveL [[-13.150,137.727,113.542],[0.15109221,-0.80885359,-0.41547485,-0.38769532],[-1,0,0,0],[9E+09,9E+09,9E+09,9E+09,9E+09,9E+09]],[16.67,500,5000,1000],z1,Weldgun \WObj:=WeldingReference;
		MoveL [[-14.061,138.456,113.433],[0.14174256,-0.81772465,-0.39285266,-0.39610886],[-1,0,0,0],[9E+09,9E+09,9E+09,9E+09,9E+09,9E+09]],[16.67,500,5000,1000],z1,Weldgun \WObj:=WeldingReference;
		MoveL [[-14.932,139.236,113.322],[0.13102406,-0.82465910,-0.37283349,-0.40467919],[-1,0,0,0],[9E+09,9E+09,9E+09,9E+09,9E+09,9E+09]],[16.67,500,5000,1000],z1,Weldgun \WObj:=WeldingReference;
		MoveL [[-15.417,139.710,113.257],[0.12572329,-0.82925325,-0.35931618,-0.40917550],[-1,0,0,0],[9E+09,9E+09,9E+09,9E+09,9E+09,9E+09]],[16.67,500,5000,1000],z1,Weldgun \WObj:=WeldingReference;
		MoveL [[-15.892,140.204,113.191],[0.12198550,-0.83499702,-0.34238421,-0.41312538],[-1,0,0,0],[9E+09,9E+09,9E+09,9E+09,9E+09,9E+09]],[16.67,500,5000,1000],z1,Weldgun \WObj:=WeldingReference;
		MoveL [[-16.680,141.100,113.078],[0.11289594,-0.84212403,-0.31822338,-0.42049437],[-1,0,0,0],[9E+09,9E+09,9E+09,9E+09,9E+09,9E+09]],[16.67,500,5000,1000],z1,Weldgun \WObj:=WeldingReference;
		MoveL [[-17.416,142.038,112.967],[0.10395269,-0.84863987,-0.29380432,-0.42741459],[-1,0,0,0],[9E+09,9E+09,9E+09,9E+09,9E+09,9E+09]],[16.67,500,5000,1000],z1,Weldgun \WObj:=WeldingReference;
		MoveL [[-18.101,143.016,112.859],[0.09514807,-0.85454646,-0.26918066,-0.43386514],[-1,0,0,0],[9E+09,9E+09,9E+09,9E+09,9E+09,9E+09]],[16.67,500,5000,1000],z1,Weldgun \WObj:=WeldingReference;
		MoveL [[-18.731,144.031,112.756],[0.08647260,-0.85985479,-0.24438897,-0.43982526],[-1,0,1,0],[9E+09,9E+09,9E+09,9E+09,9E+09,9E+09]],[16.67,500,5000,1000],z1,Weldgun \WObj:=WeldingReference;
		MoveL [[-19.306,145.081,112.659],[0.07792686,-0.86457595,-0.21946800,-0.44527478],[-1,0,1,0],[9E+09,9E+09,9E+09,9E+09,9E+09,9E+09]],[16.67,500,5000,1000],z1,Weldgun \WObj:=WeldingReference;
		MoveL [[-19.824,146.161,112.569],[0.06949759,-0.86872617,-0.19443195,-0.45020122],[-1,0,1,0],[9E+09,9E+09,9E+09,9E+09,9E+09,9E+09]],[16.67,500,5000,1000],z1,Weldgun \WObj:=WeldingReference;
		MoveL [[-20.284,147.270,112.487],[0.06115910,-0.87231524,-0.16933251,-0.45459013],[-1,0,1,0],[9E+09,9E+09,9E+09,9E+09,9E+09,9E+09]],[16.67,500,5000,1000],z1,Weldgun \WObj:=WeldingReference;
		MoveL [[-20.685,148.403,112.414],[0.05292637,-0.87536045,-0.14417663,-0.45842773],[-1,0,1,0],[9E+09,9E+09,9E+09,9E+09,9E+09,9E+09]],[16.67,500,5000,1000],z1,Weldgun \WObj:=WeldingReference;
		MoveL [[-21.026,149.557,112.351],[0.04478259,-0.87787936,-0.11895843,-0.46170471],[-1,0,1,0],[9E+09,9E+09,9E+09,9E+09,9E+09,9E+09]],[16.67,500,5000,1000],z1,Weldgun \WObj:=WeldingReference;
		MoveL [[-21.307,150.732,112.298],[0.03668848,-0.87988914,-0.09360872,-0.46442057],[-1,0,1,0],[9E+09,9E+09,9E+09,9E+09,9E+09,9E+09]],[16.67,500,5000,1000],z1,Weldgun \WObj:=WeldingReference;
		MoveL [[-21.528,151.930,112.256],[0.02856986,-0.88139032,-0.06814633,-0.46657362],[-1,0,1,0],[9E+09,9E+09,9E+09,9E+09,9E+09,9E+09]],[16.67,500,5000,1000],z1,Weldgun \WObj:=WeldingReference;
		MoveL [[-21.686,153.139,112.225],[0.02048892,-0.88238735,-0.04267608,-0.46813623],[-1,0,1,0],[9E+09,9E+09,9E+09,9E+09,9E+09,9E+09]],[16.67,500,5000,1000],z1,Weldgun \WObj:=WeldingReference;
		MoveL [[-21.782,154.355,112.207],[0.01243893,-0.88288728,-0.01720659,-0.46910473],[-1,0,1,0],[9E+09,9E+09,9E+09,9E+09,9E+09,9E+09]],[16.67,500,5000,1000],z1,Weldgun \WObj:=WeldingReference;
		MoveL [[-21.813,155.575,112.201],[0.00000000,0.88293325,0.00000000,0.46949853],[-1,0,1,0],[9E+09,9E+09,9E+09,9E+09,9E+09,9E+09]],[16.67,500,5000,1000],z1,Weldgun \WObj:=WeldingReference;
		MoveL [[-21.813,184.150,112.201],[0.00586319,0.88286421,0.01101837,0.46946246],[-1,0,1,0],[9E+09,9E+09,9E+09,9E+09,9E+09,9E+09]],[16.67,500,5000,1000],z1,Weldgun \WObj:=WeldingReference;
		MoveL [[-21.814,185.241,112.169],[0.03165533,0.88236559,0.02554723,0.46880299],[-1,0,1,0],[9E+09,9E+09,9E+09,9E+09,9E+09,9E+09]],[16.67,500,5000,1000],z1,Weldgun \WObj:=WeldingReference;
		MoveL [[-21.818,186.329,112.072],[0.05742808,0.88123291,0.04001861,0.46747095],[-1,0,1,0],[9E+09,9E+09,9E+09,9E+09,9E+09,9E+09]],[16.67,500,5000,1000],z1,Weldgun \WObj:=WeldingReference;
		MoveL [[-21.823,187.410,111.912],[0.08316160,0.87946762,0.05439385,0.46546982],[-1,0,1,0],[9E+09,9E+09,9E+09,9E+09,9E+09,9E+09]],[16.67,500,5000,1000],z1,Weldgun \WObj:=WeldingReference;
		MoveL [[-21.831,188.481,111.689],[0.10883995,0.87707132,0.06862859,0.46280653],[-1,0,1,0],[9E+09,9E+09,9E+09,9E+09,9E+09,9E+09]],[16.67,500,5000,1000],z1,Weldgun \WObj:=WeldingReference;
		MoveL [[-21.841,189.538,111.403],[0.13444877,0.87404675,0.08268225,0.45948824],[-1,0,1,0],[9E+09,9E+09,9E+09,9E+09,9E+09,9E+09]],[16.67,500,5000,1000],z1,Weldgun \WObj:=WeldingReference;
		MoveL [[-21.854,190.577,111.055],[0.15998221,0.87039388,0.09652688,0.45552470],[-1,0,1,0],[9E+09,9E+09,9E+09,9E+09,9E+09,9E+09]],[16.67,500,5000,1000],z1,Weldgun \WObj:=WeldingReference;
		MoveL [[-21.868,191.597,110.645],[0.18540893,0.86611896,0.11010253,0.45093115],[-1,0,1,0],[9E+09,9E+09,9E+09,9E+09,9E+09,9E+09]],[16.67,500,5000,1000],z1,Weldgun \WObj:=WeldingReference;
		MoveL [[-21.884,192.593,110.176],[0.21074379,0.86121856,0.12338373,0.44571976],[-1,0,1,0],[9E+09,9E+09,9E+09,9E+09,9E+09,9E+09]],[16.67,500,5000,1000],z1,Weldgun \WObj:=WeldingReference;
		MoveL [[-21.901,193.562,109.648],[0.23595306,0.85569953,0.13633443,0.43990612],[-1,0,1,0],[9E+09,9E+09,9E+09,9E+09,9E+09,9E+09]],[16.67,500,5000,1000],z1,Weldgun \WObj:=WeldingReference;
		MoveL [[-21.921,194.501,109.063],[0.25867767,0.85035795,0.14428354,0.43492469],[-1,0,1,0],[9E+09,9E+09,9E+09,9E+09,9E+09,9E+09]],[16.67,500,5000,1000],z1,Weldgun \WObj:=WeldingReference;
		MoveL [[-21.932,195.003,108.718],[0.27239128,0.84676957,0.15098755,0.43126215],[-1,0,1,0],[9E+09,9E+09,9E+09,9E+09,9E+09,9E+09]],[16.67,500,5000,1000],z1,Weldgun \WObj:=WeldingReference;
		MoveL [[-21.944,195.488,108.361],[0.28874100,0.84197226,0.16311317,0.42556485],[-1,0,1,0],[9E+09,9E+09,9E+09,9E+09,9E+09,9E+09]],[16.67,500,5000,1000],z1,Weldgun \WObj:=WeldingReference;
		MoveL [[-21.968,196.435,107.592],[0.31535543,0.83400435,0.17484577,0.41763220],[-1,0,1,0],[9E+09,9E+09,9E+09,9E+09,9E+09,9E+09]],[16.67,500,5000,1000],z1,Weldgun \WObj:=WeldingReference;
		MoveL [[-21.991,197.253,106.841],[0.33979058,0.82596253,0.18591056,0.40959191],[-1,0,1,0],[9E+09,9E+09,9E+09,9E+09,9E+09,9E+09]],[16.67,500,5000,1000],z1,Weldgun \WObj:=WeldingReference;
		MoveL [[-22.014,198.028,106.041],[0.36404560,0.81731975,0.19643477,0.40108927],[-1,0,1,0],[9E+09,9E+09,9E+09,9E+09,9E+09,9E+09]],[16.67,500,5000,1000],z1,Weldgun \WObj:=WeldingReference;
		MoveL [[-22.038,198.757,105.197],[0.38806259,0.80809146,0.20641310,0.39215973],[-1,0,1,0],[9E+09,9E+09,9E+09,9E+09,9E+09,9E+09]],[16.67,500,5000,1000],z1,Weldgun \WObj:=WeldingReference;
		MoveL [[-22.062,199.440,104.308],[0.41187949,0.79826576,0.21579762,0.38282953],[-1,0,1,0],[9E+09,9E+09,9E+09,9E+09,9E+09,9E+09]],[16.67,500,5000,1000],z1,Weldgun \WObj:=WeldingReference;
		MoveL [[-22.085,200.070,103.381],[0.43543412,0.78786159,0.22456360,0.37315203],[-1,0,1,0],[9E+09,9E+09,9E+09,9E+09,9E+09,9E+09]],[16.67,500,5000,1000],z1,Weldgun \WObj:=WeldingReference;
		MoveL [[-22.108,200.648,102.418],[0.45871624,0.77688323,0.23268585,0.36316546],[-1,0,1,0],[9E+09,9E+09,9E+09,9E+09,9E+09,9E+09]],[16.67,500,5000,1000],z1,Weldgun \WObj:=WeldingReference;
		MoveL [[-22.130,201.171,101.422],[0.48171990,0.76532819,0.24017170,0.35289694],[-1,0,1,0],[9E+09,9E+09,9E+09,9E+09,9E+09,9E+09]],[16.67,500,5000,1000],z1,Weldgun \WObj:=WeldingReference;
		MoveL [[-22.151,201.637,100.396],[0.50444957,0.75318944,0.24698755,0.34239371],[-1,0,1,0],[9E+09,9E+09,9E+09,9E+09,9E+09,9E+09]],[16.67,500,5000,1000],z1,Weldgun \WObj:=WeldingReference;
		MoveL [[-22.169,202.045,99.343],[0.52689169,0.74046558,0.25314512,0.33168271],[-1,0,1,0],[9E+09,9E+09,9E+09,9E+09,9E+09,9E+09]],[16.67,500,5000,1000],z1,Weldgun \WObj:=WeldingReference;
		MoveL [[-22.186,202.393,98.266],[0.54599414,0.72955538,0.25172687,0.32599528],[-1,0,1,0],[9E+09,9E+09,9E+09,9E+09,9E+09,9E+09]],[16.67,500,5000,1000],z1,Weldgun \WObj:=WeldingReference;
		MoveL [[-22.176,202.643,97.334],[0.57084032,0.71283198,0.23939194,0.32970198],[-1,0,1,0],[9E+09,9E+09,9E+09,9E+09,9E+09,9E+09]],[16.67,500,5000,1000],z1,Weldgun \WObj:=WeldingReference;
		MoveL [[-22.147,202.775,96.757],[0.58584689,0.70188649,0.23158017,0.33242954],[-1,0,1,0],[9E+09,9E+09,9E+09,9E+09,9E+09,9E+09]],[16.67,500,5000,1000],z1,Weldgun \WObj:=WeldingReference;
		MoveL [[-22.099,202.892,96.163],[0.60136158,0.68988462,0.22430189,0.33483148],[-1,0,1,0],[9E+09,9E+09,9E+09,9E+09,9E+09,9E+09]],[16.67,500,5000,1000],z1,Weldgun \WObj:=WeldingReference;
		MoveL [[-21.988,203.039,95.230],[0.62490710,0.67020270,0.21276965,0.33918804],[-1,0,1,0],[9E+09,9E+09,9E+09,9E+09,9E+09,9E+09]],[16.67,500,5000,1000],z1,Weldgun \WObj:=WeldingReference;
		MoveL [[-21.835,203.138,94.305],[0.64763111,0.64941747,0.20197666,0.34356414],[-1,0,1,0],[9E+09,9E+09,9E+09,9E+09,9E+09,9E+09]],[16.67,500,5000,1000],z1,Weldgun \WObj:=WeldingReference;
		MoveL [[-21.639,203.192,93.372],[0.66881390,0.62786082,0.19023049,0.34970147],[-1,0,1,0],[9E+09,9E+09,9E+09,9E+09,9E+09,9E+09]],[16.67,500,5000,1000],z1,Weldgun \WObj:=WeldingReference;
		MoveL [[-21.328,203.201,92.188],[0.68119986,0.61013554,0.16880665,0.36770325],[-1,0,2,0],[9E+09,9E+09,9E+09,9E+09,9E+09,9E+09]],[16.67,500,5000,1000],z1,Weldgun \WObj:=WeldingReference;
		MoveL [[-20.918,203.201,90.925],[0.68593960,0.59887738,0.14838059,0.38576670],[-1,0,2,0],[9E+09,9E+09,9E+09,9E+09,9E+09,9E+09]],[16.67,500,5000,1000],z1,Weldgun \WObj:=WeldingReference;
		MoveL [[-20.432,203.201,89.689],[0.69006493,0.58708440,0.12781765,0.40349095],[-1,0,2,0],[9E+09,9E+09,9E+09,9E+09,9E+09,9E+09]],[16.67,500,5000,1000],z1,Weldgun \WObj:=WeldingReference;
		MoveL [[-19.874,203.201,88.484],[0.69357798,0.57476662,0.10714562,0.42084764],[-1,0,2,0],[9E+09,9E+09,9E+09,9E+09,9E+09,9E+09]],[16.67,500,5000,1000],z1,Weldgun \WObj:=WeldingReference;
		MoveL [[-19.245,203.201,87.315],[0.69646838,0.56193667,0.08637475,0.43783375],[-1,0,2,0],[9E+09,9E+09,9E+09,9E+09,9E+09,9E+09]],[16.67,500,5000,1000],z1,Weldgun \WObj:=WeldingReference;
		MoveL [[-18.547,203.201,86.185],[0.69873897,0.54860461,0.06552875,0.45442581],[-1,0,2,0],[9E+09,9E+09,9E+09,9E+09,9E+09,9E+09]],[16.67,500,5000,1000],z1,Weldgun \WObj:=WeldingReference;
		MoveL [[-17.783,203.201,85.099],[0.70038377,0.53478284,0.04462157,0.47061535],[-1,0,2,0],[9E+09,9E+09,9E+09,9E+09,9E+09,9E+09]],[16.67,500,5000,1000],z1,Weldgun \WObj:=WeldingReference;
		MoveL [[-16.955,203.201,84.061],[0.70140586,0.52048344,0.02367788,0.48638068],[-1,0,2,0],[9E+09,9E+09,9E+09,9E+09,9E+09,9E+09]],[16.67,500,5000,1000],z1,Weldgun \WObj:=WeldingReference;
		MoveL [[-16.067,203.201,83.074],[0.70179746,0.50571955,0.00270884,0.50171778],[-1,0,2,0],[9E+09,9E+09,9E+09,9E+09,9E+09,9E+09]],[16.67,500,5000,1000],z1,Weldgun \WObj:=WeldingReference;
		MoveL [[-15.121,203.201,82.142],[0.70241235,0.49053286,-0.01745484,0.51545100],[-1,0,2,0],[9E+09,9E+09,9E+09,9E+09,9E+09,9E+09]],[16.67,500,5000,1000],z1,Weldgun \WObj:=WeldingReference;
		MoveL [[-14.280,203.201,81.399],[0.70171587,0.47736356,-0.03520854,0.52771131],[-1,0,2,0],[9E+09,9E+09,9E+09,9E+09,9E+09,9E+09]],[16.67,500,5000,1000],z1,Weldgun \WObj:=WeldingReference;
		MoveL [[-13.397,203.201,80.696],[0.70030181,0.46376974,-0.05328194,0.54005188],[-1,0,2,0],[9E+09,9E+09,9E+09,9E+09,9E+09,9E+09]],[16.67,500,5000,1000],z1,Weldgun \WObj:=WeldingReference;
		MoveL [[-12.422,203.201,79.999],[0.69860821,0.44904066,-0.07214449,0.55236241],[-1,0,2,0],[9E+09,9E+09,9E+09,9E+09,9E+09,9E+09]],[16.67,500,5000,1000],z1,Weldgun \WObj:=WeldingReference;
		MoveL [[-11.410,203.201,79.357],[0.69640996,0.43398715,-0.09095072,0.56426614],[-1,0,2,0],[9E+09,9E+09,9E+09,9E+09,9E+09,9E+09]],[16.67,500,5000,1000],z1,Weldgun \WObj:=WeldingReference;
		MoveL [[-10.366,203.201,78.769],[0.69370517,0.41861709,-0.10969168,0.57576089],[-1,0,2,0],[9E+09,9E+09,9E+09,9E+09,9E+09,9E+09]],[16.67,500,5000,1000],z1,Weldgun \WObj:=WeldingReference;
		MoveL [[-9.292,203.201,78.239],[0.69049479,0.40294288,-0.12835522,0.58683806],[-1,0,2,0],[9E+09,9E+09,9E+09,9E+09,9E+09,9E+09]],[16.67,500,5000,1000],z1,Weldgun \WObj:=WeldingReference;
		MoveL [[-8.190,203.201,77.768],[0.68678461,0.38697602,-0.14692248,0.59748661],[-1,0,2,0],[9E+09,9E+09,9E+09,9E+09,9E+09,9E+09]],[16.67,500,5000,1000],z1,Weldgun \WObj:=WeldingReference;
		MoveL [[-7.065,203.201,77.356],[0.68257350,0.37072825,-0.16538378,0.60770239],[-1,0,2,0],[9E+09,9E+09,9E+09,9E+09,9E+09,9E+09]],[16.67,500,5000,1000],z1,Weldgun \WObj:=WeldingReference;
		MoveL [[-5.919,203.201,77.006],[0.67786869,0.35421122,-0.18372425,0.61747376],[-1,0,2,0],[9E+09,9E+09,9E+09,9E+09,9E+09,9E+09]],[16.67,500,5000,1000],z1,Weldgun \WObj:=WeldingReference;
		MoveL [[-4.756,203.201,76.719],[0.67266523,0.33743479,-0.20193424,0.62680285],[-1,0,2,0],[9E+09,9E+09,9E+09,9E+09,9E+09,9E+09]],[16.67,500,5000,1000],z1,Weldgun \WObj:=WeldingReference;
		MoveL [[-3.579,203.201,76.494],[0.66698095,0.32041557,-0.21999343,0.63566749],[-1,0,2,0],[9E+09,9E+09,9E+09,9E+09,9E+09,9E+09]],[16.67,500,5000,1000],z1,Weldgun \WObj:=WeldingReference;
		MoveL [[-2.392,203.201,76.333],[0.66080513,0.30316129,-0.23789569,0.64407721],[-1,0,2,0],[9E+09,9E+09,9E+09,9E+09,9E+09,9E+09]],[16.67,500,5000,1000],z1,Weldgun \WObj:=WeldingReference;
		MoveL [[-1.198,203.201,76.236],[0.65415296,0.28568786,-0.25562294,0.65201478],[-1,0,2,0],[9E+09,9E+09,9E+09,9E+09,9E+09,9E+09]],[16.67,500,5000,1000],z1,Weldgun \WObj:=WeldingReference;
		MoveL [[0.000,203.201,76.204],[0.64702338,0.26800578,-0.27316590,0.65948013],[-1,0,2,0],[9E+09,9E+09,9E+09,9E+09,9E+09,9E+09]],[16.67,500,5000,1000],z1,Weldgun \WObj:=WeldingReference;
		MoveL [[1.198,203.201,76.236],[0.63942538,0.25012984,-0.29050880,0.66646446],[-1,0,2,0],[9E+09,9E+09,9E+09,9E+09,9E+09,9E+09]],[16.67,500,5000,1000],z1,Weldgun \WObj:=WeldingReference;
		MoveL [[2.392,203.201,76.333],[0.63135831,0.23207101,-0.30764287,0.67296775],[-1,0,2,0],[9E+09,9E+09,9E+09,9E+09,9E+09,9E+09]],[16.67,500,5000,1000],z1,Weldgun \WObj:=WeldingReference;
		MoveL [[3.579,203.201,76.494],[0.62284124,0.21384548,-0.32455097,0.67897391],[-1,0,2,0],[9E+09,9E+09,9E+09,9E+09,9E+09,9E+09]],[16.67,500,5000,1000],z1,Weldgun \WObj:=WeldingReference;
		MoveL [[4.756,203.201,76.719],[0.61386100,0.19546092,-0.34122510,0.68449626],[-1,0,3,0],[9E+09,9E+09,9E+09,9E+09,9E+09,9E+09]],[16.67,500,5000,1000],z1,Weldgun \WObj:=WeldingReference;
		MoveL [[5.919,203.201,77.006],[0.60443803,0.17693903,-0.35764863,0.68951774],[-1,-1,3,0],[9E+09,9E+09,9E+09,9E+09,9E+09,9E+09]],[16.67,500,5000,1000],z1,Weldgun \WObj:=WeldingReference;
		MoveL [[7.065,203.201,77.356],[0.59457495,0.15828650,-0.37381353,0.69403851],[-1,-1,3,0],[9E+09,9E+09,9E+09,9E+09,9E+09,9E+09]],[16.67,500,5000,1000],z1,Weldgun \WObj:=WeldingReference;
		MoveL [[8.190,203.201,77.768],[0.58428714,0.13951697,-0.38970780,0.69804827],[-1,-1,3,0],[9E+09,9E+09,9E+09,9E+09,9E+09,9E+09]],[16.67,500,5000,1000],z1,Weldgun \WObj:=WeldingReference;
		MoveL [[9.292,203.201,78.239],[0.57356464,0.12064858,-0.40531712,0.70155938],[-1,-1,3,0],[9E+09,9E+09,9E+09,9E+09,9E+09,9E+09]],[16.67,500,5000,1000],z1,Weldgun \WObj:=WeldingReference;
		MoveL [[10.366,203.201,78.769],[0.56242858,0.10169157,-0.42063240,0.70455753],[-1,-1,3,0],[9E+09,9E+09,9E+09,9E+09,9E+09,9E+09]],[16.67,500,5000,1000],z1,Weldgun \WObj:=WeldingReference;
		MoveL [[11.410,203.201,79.357],[0.55088743,0.08266025,-0.43564212,0.70704050],[-1,-1,3,0],[9E+09,9E+09,9E+09,9E+09,9E+09,9E+09]],[16.67,500,5000,1000],z1,Weldgun \WObj:=WeldingReference;
		MoveL [[12.422,203.201,79.999],[0.53893865,0.06356691,-0.45033561,0.70901496],[-1,-1,3,0],[9E+09,9E+09,9E+09,9E+09,9E+09,9E+09]],[16.67,500,5000,1000],z1,Weldgun \WObj:=WeldingReference;
		MoveL [[13.397,203.201,80.696],[0.52738231,0.04493855,-0.46465215,0.70989210],[-1,-1,3,0],[9E+09,9E+09,9E+09,9E+09,9E+09,9E+09]],[16.67,500,5000,1000],z1,Weldgun \WObj:=WeldingReference;
		MoveL [[14.227,203.201,81.355],[0.51609769,0.02795371,-0.47710917,0.71079435],[-1,-1,3,0],[9E+09,9E+09,9E+09,9E+09,9E+09,9E+09]],[16.67,500,5000,1000],z1,Weldgun \WObj:=WeldingReference;
		MoveL [[15.031,203.201,82.059],[0.50301183,0.00984587,-0.48939955,0.71229926],[-1,-1,3,0],[9E+09,9E+09,9E+09,9E+09,9E+09,9E+09]],[16.67,500,5000,1000],z1,Weldgun \WObj:=WeldingReference;
		MoveL [[15.982,203.201,82.986],[0.48816215,-0.01143852,-0.50420960,0.71227772],[-1,-1,3,0],[9E+09,9E+09,9E+09,9E+09,9E+09,9E+09]],[16.67,500,5000,1000],z1,Weldgun \WObj:=WeldingReference;
		MoveL [[16.876,203.201,83.968],[0.47288185,-0.03271617,-0.51856953,0.71161650],[-1,-1,3,0],[9E+09,9E+09,9E+09,9E+09,9E+09,9E+09]],[16.67,500,5000,1000],z1,Weldgun \WObj:=WeldingReference;
		MoveL [[17.709,203.201,85.002],[0.45717321,-0.05396142,-0.53246628,0.71032421],[-1,-1,3,0],[9E+09,9E+09,9E+09,9E+09,9E+09,9E+09]],[16.67,500,5000,1000],z1,Weldgun \WObj:=WeldingReference;
		MoveL [[18.479,203.201,86.084],[0.44106469,-0.07516210,-0.54588738,0.70839224],[-1,-1,3,0],[9E+09,9E+09,9E+09,9E+09,9E+09,9E+09]],[16.67,500,5000,1000],z1,Weldgun \WObj:=WeldingReference;
		MoveL [[19.183,203.201,87.209],[0.42455597,-0.09629090,-0.55882195,0.70583165],[-1,-1,3,0],[9E+09,9E+09,9E+09,9E+09,9E+09,9E+09]],[16.67,500,5000,1000],z1,Weldgun \WObj:=WeldingReference;
		MoveL [[19.819,203.201,88.375],[0.40766840,-0.11733640,-0.57125642,0.70264127],[-1,-1,3,0],[9E+09,9E+09,9E+09,9E+09,9E+09,9E+09]],[16.67,500,5000,1000],z1,Weldgun \WObj:=WeldingReference;
		MoveL [[20.384,203.201,89.577],[0.39042413,-0.13827833,-0.58318156,0.69881855],[-1,-1,3,0],[9E+09,9E+09,9E+09,9E+09,9E+09,9E+09]],[16.67,500,5000,1000],z1,Weldgun \WObj:=WeldingReference;
		MoveL [[20.876,203.201,90.810],[0.37282190,-0.15909440,-0.59458602,0.69437762],[-1,-1,3,0],[9E+09,9E+09,9E+09,9E+09,9E+09,9E+09]],[16.67,500,5000,1000],z1,Weldgun \WObj:=WeldingReference;
		MoveL [[21.294,203.201,92.070],[0.35656803,-0.17829782,-0.60589441,0.68844832],[-1,-1,3,0],[9E+09,9E+09,9E+09,9E+09,9E+09,9E+09]],[16.67,500,5000,1000],z1,Weldgun \WObj:=WeldingReference;
		MoveL [[21.625,203.194,93.309],[0.35007295,-0.18951337,-0.62634225,0.67024548],[-1,0,3,0],[9E+09,9E+09,9E+09,9E+09,9E+09,9E+09]],[16.67,500,5000,1000],z1,Weldgun \WObj:=WeldingReference;
		MoveL [[21.830,203.141,94.271],[0.34515387,-0.20017116,-0.64908984,0.64767483],[-1,0,3,0],[9E+09,9E+09,9E+09,9E+09,9E+09,9E+09]],[16.67,500,5000,1000],z1,Weldgun \WObj:=WeldingReference;
		MoveL [[21.989,203.039,95.230],[0.34026254,-0.21161558,-0.67056821,0.62432246],[-1,0,3,0],[9E+09,9E+09,9E+09,9E+09,9E+09,9E+09]],[16.67,500,5000,1000],z1,Weldgun \WObj:=WeldingReference;
		MoveL [[22.102,202.887,96.188],[0.33512237,-0.22415853,-0.69055437,0.60048365],[-1,0,3,0],[9E+09,9E+09,9E+09,9E+09,9E+09,9E+09]],[16.67,500,5000,1000],z1,Weldgun \WObj:=WeldingReference;
		MoveL [[22.147,202.775,96.757],[0.33301213,-0.23087937,-0.70211759,0.58551562],[-1,0,3,0],[9E+09,9E+09,9E+09,9E+09,9E+09,9E+09]],[16.67,500,5000,1000],z1,Weldgun \WObj:=WeldingReference;
		MoveL [[22.176,202.645,97.326],[0.33038784,-0.23847681,-0.71294636,0.57068395],[-1,0,3,0],[9E+09,9E+09,9E+09,9E+09,9E+09,9E+09]],[16.67,500,5000,1000],z1,Weldgun \WObj:=WeldingReference;
		MoveL [[22.186,202.393,98.266],[0.33198844,-0.24367277,-0.73228810,0.54236648],[-1,0,3,0],[9E+09,9E+09,9E+09,9E+09,9E+09,9E+09]],[16.67,500,5000,1000],z1,Weldgun \WObj:=WeldingReference;
		MoveL [[22.169,202.045,99.343],[0.34259161,-0.23765753,-0.74557852,0.51986783],[-1,0,3,0],[9E+09,9E+09,9E+09,9E+09,9E+09,9E+09]],[16.67,500,5000,1000],z1,Weldgun \WObj:=WeldingReference;
		MoveL [[22.151,201.637,100.396],[0.35299929,-0.23097809,-0.75825608,0.49707981],[-1,0,3,0],[9E+09,9E+09,9E+09,9E+09,9E+09,9E+09]],[16.67,500,5000,1000],z1,Weldgun \WObj:=WeldingReference;
		MoveL [[22.130,201.171,101.422],[0.36319068,-0.22363105,-0.77032123,0.47401149],[-1,0,3,0],[9E+09,9E+09,9E+09,9E+09,9E+09,9E+09]],[16.67,500,5000,1000],z1,Weldgun \WObj:=WeldingReference;
		MoveL [[22.108,200.648,102.418],[0.37311180,-0.21564402,-0.78178523,0.45066295],[-1,0,3,0],[9E+09,9E+09,9E+09,9E+09,9E+09,9E+09]],[16.67,500,5000,1000],z1,Weldgun \WObj:=WeldingReference;
		MoveL [[22.085,200.070,103.381],[0.38273018,-0.20700438,-0.79265820,0.42703603],[-1,0,3,0],[9E+09,9E+09,9E+09,9E+09,9E+09,9E+09]],[16.67,500,5000,1000],z1,Weldgun \WObj:=WeldingReference;
		MoveL [[22.062,199.440,104.308],[0.39201635,-0.19774541,-0.80292628,0.40314926],[-1,0,3,0],[9E+09,9E+09,9E+09,9E+09,9E+09,9E+09]],[16.67,500,5000,1000],z1,Weldgun \WObj:=WeldingReference;
		MoveL [[22.038,198.757,105.197],[0.40091142,-0.18791559,-0.81259460,0.37900895],[-1,0,3,0],[9E+09,9E+09,9E+09,9E+09,9E+09,9E+09]],[16.67,500,5000,1000],z1,Weldgun \WObj:=WeldingReference;
		MoveL [[22.014,198.028,106.041],[0.40939227,-0.17750857,-0.82163762,0.35468338],[-1,0,3,0],[9E+09,9E+09,9E+09,9E+09,9E+09,9E+09]],[16.67,500,5000,1000],z1,Weldgun \WObj:=WeldingReference;
		MoveL [[21.991,197.253,106.841],[0.41741536,-0.16657481,-0.83007727,0.33013479],[-1,0,3,0],[9E+09,9E+09,9E+09,9E+09,9E+09,9E+09]],[16.67,500,5000,1000],z1,Weldgun \WObj:=WeldingReference;
		MoveL [[21.968,196.435,107.592],[0.42349774,-0.15911270,-0.83714654,0.30743859],[-1,0,3,0],[9E+09,9E+09,9E+09,9E+09,9E+09,9E+09]],[16.67,500,5000,1000],z1,Weldgun \WObj:=WeldingReference;
		MoveL [[21.954,195.926,108.018],[0.42781750,-0.15211072,-0.84155462,0.29260952],[-1,0,3,0],[9E+09,9E+09,9E+09,9E+09,9E+09,9E+09]],[16.67,500,5000,1000],z1,Weldgun \WObj:=WeldingReference;
		MoveL [[21.942,195.407,108.422],[0.43328375,-0.14083305,-0.84642114,0.27568549],[-1,0,3,0],[9E+09,9E+09,9E+09,9E+09,9E+09,9E+09]],[16.67,500,5000,1000],z1,Weldgun \WObj:=WeldingReference;
		MoveL [[21.921,194.501,109.063],[0.43968334,-0.12836672,-0.85290498,0.25050677],[-1,0,3,0],[9E+09,9E+09,9E+09,9E+09,9E+09,9E+09]],[16.67,500,5000,1000],z1,Weldgun \WObj:=WeldingReference;
		MoveL [[21.901,193.562,109.648],[0.44550693,-0.11551765,-0.85875730,0.22520025],[-1,0,3,0],[9E+09,9E+09,9E+09,9E+09,9E+09,9E+09]],[16.67,500,5000,1000],z1,Weldgun \WObj:=WeldingReference;
		MoveL [[21.884,192.593,110.176],[0.45073466,-0.10231387,-0.86397472,0.19979446],[-1,0,3,0],[9E+09,9E+09,9E+09,9E+09,9E+09,9E+09]],[16.67,500,5000,1000],z1,Weldgun \WObj:=WeldingReference;
		MoveL [[21.868,191.597,110.645],[0.45534645,-0.08881484,-0.86855913,0.17428875],[-1,0,3,0],[9E+09,9E+09,9E+09,9E+09,9E+09,9E+09]],[16.67,500,5000,1000],z1,Weldgun \WObj:=WeldingReference;
		MoveL [[21.854,190.577,111.055],[0.45933182,-0.07503473,-0.87251063,0.14869185],[-1,0,3,0],[9E+09,9E+09,9E+09,9E+09,9E+09,9E+09]],[16.67,500,5000,1000],z1,Weldgun \WObj:=WeldingReference;
		MoveL [[21.841,189.538,111.403],[0.46267440,-0.06102668,-0.87582540,0.12303665],[-1,0,3,0],[9E+09,9E+09,9E+09,9E+09,9E+09,9E+09]],[16.67,500,5000,1000],z1,Weldgun \WObj:=WeldingReference;
		MoveL [[21.831,188.481,111.689],[0.46536551,-0.04683904,-0.87850496,0.09731438],[-1,0,3,0],[9E+09,9E+09,9E+09,9E+09,9E+09,9E+09]],[16.67,500,5000,1000],z1,Weldgun \WObj:=WeldingReference;
		MoveL [[21.823,187.410,111.912],[0.46739520,-0.03249057,-0.88054870,0.07155476],[-1,0,3,0],[9E+09,9E+09,9E+09,9E+09,9E+09,9E+09]],[16.67,500,5000,1000],z1,Weldgun \WObj:=WeldingReference;
		MoveL [[21.818,186.329,112.072],[0.46875684,-0.01804249,-0.88195674,0.04575809],[-1,0,3,0],[9E+09,9E+09,9E+09,9E+09,9E+09,9E+09]],[16.67,500,5000,1000],z1,Weldgun \WObj:=WeldingReference;
		MoveL [[21.814,185.241,112.169],[0.46944730,-0.00352434,-0.88272803,0.01995068],[-1,0,3,0],[9E+09,9E+09,9E+09,9E+09,9E+09,9E+09]],[16.67,500,5000,1000],z1,Weldgun \WObj:=WeldingReference;
		MoveL [[21.813,184.150,112.201],[0.46949853,-0.00000000,-0.88293325,0.00000000],[-1,0,3,0],[9E+09,9E+09,9E+09,9E+09,9E+09,9E+09]],[16.67,500,5000,1000],z1,Weldgun \WObj:=WeldingReference;
		MoveL [[21.813,169.863,112.201],[0.46949853,0.00000000,-0.88293325,-0.00000000],[-1,0,3,0],[9E+09,9E+09,9E+09,9E+09,9E+09,9E+09]],[16.67,500,5000,1000],z1,Weldgun \WObj:=WeldingReference;
		GunOff;
		MoveL [[21.813,169.863,112.201],[0.46949853,0.00000000,-0.88293325,-0.00000000],[-1,0,3,0],[9E+09,9E+09,9E+09,9E+09,9E+09,9E+09]],v1000,z1,Weldgun \WObj:=WeldingReference;
		MoveL [[104.720,169.863,168.115],[0.46905216,-0.03851172,-0.88209262,0.02048227],[-1,0,3,0],[9E+09,9E+09,9E+09,9E+09,9E+09,9E+09]],v1000,z1,Weldgun \WObj:=WeldingReference;
	ENDPROC

	PROC Main()
		ConfJ \On;
		ConfL \Off;
		! Program generated by VerticalBot Studio for ABB IRB 2600-12/1.65 on 25/10/2026 12:00:00
		! Using nominal kinematics.
		GoHome;
		Weld1;
		GoHome;
		Weld2;
		GoHome;
		Weld3;
		GoHome;
	ENDPROC

ENDMODULE
